(*
	FIFO queue that owns every FB_LogRecord pointer it contains. push drops the
	oldest owned records when the bound is reached. The bound is maxCount, but
	never more than TcOtlp_GVL.MAX_LOOP_COUNT: a maxCount of zero, or one above
	that limit, is held to MAX_LOOP_COUNT so that free always reaches the end.
	pop transfers ownership back to the caller. transferTo moves allocated
	nodes between queue owners without copying records.
*)
FUNCTION_BLOCK FB_LogRecordQueue
VAR
	_head: POINTER TO ST_LinkedListNode;
	_tail: POINTER TO ST_LinkedListNode;
	_cursor: POINTER TO ST_LinkedListNode;
END_VAR
VAR_OUTPUT
	count: UDINT;
	maxCount: UDINT;
	droppedCount: UDINT;
END_VAR

(* The enforced bound: maxCount, held to MAX_LOOP_COUNT when it is zero or larger. *)
METHOD _capacity : UDINT
IF THIS^.maxCount = 0 OR THIS^.maxCount > TcOtlp_GVL.MAX_LOOP_COUNT THEN
	_capacity := TcOtlp_GVL.MAX_LOOP_COUNT;
ELSE
	_capacity := THIS^.maxCount;
END_IF
END_METHOD

METHOD FB_Exit : BOOL
VAR_INPUT
	bInCopyCode: BOOL;
END_VAR
IF NOT bInCopyCode THEN
	THIS^.free();
END_IF
END_METHOD

METHOD FB_Init : BOOL
VAR_INPUT
	bInitRetains: BOOL;
	bInCopyCode: BOOL;
	maxCount: UDINT := 0;
END_VAR
THIS^.maxCount := maxCount;
END_METHOD

(*
	Releases every owned record. push holds count to MAX_LOOP_COUNT, so the loop
	always reaches the end. If it ever stops early, the unreleased nodes stay in
	the queue and free returns FALSE, so a later call can finish the job.
*)
METHOD free : BOOL
VAR
	_idx: UDINT;
	_node: POINTER TO ST_LinkedListNode;
	_record: POINTER TO FB_LogRecord;
END_VAR
FOR _idx := 0 TO TcOtlp_GVL.MAX_LOOP_COUNT DO
	IF THIS^._head = 0 THEN
		EXIT;
	END_IF

	_node := THIS^._head;
	THIS^._head := _node^.nxt;
	IF _node^.val <> 0 THEN
		_record := _node^.val;
		_node^.val := 0;
		_record^.delete(pSelf:=_record);
	END_IF
	__DELETE(_node);
	IF THIS^.count > 0 THEN
		THIS^.count := THIS^.count - 1;
	END_IF
END_FOR

THIS^._cursor := THIS^._head;
IF THIS^._head = 0 THEN
	THIS^._tail := 0;
	THIS^.count := 0;
END_IF
free := THIS^._head = 0;
END_METHOD

METHOD next : POINTER TO FB_LogRecord
next := 0;

IF THIS^._cursor <> 0 THEN
	next := THIS^._cursor^.val;
	THIS^._cursor := THIS^._cursor^.nxt;
END_IF
END_METHOD

METHOD pop : BOOL
VAR_IN_OUT
	pValue: POINTER TO FB_LogRecord;
END_VAR
VAR_OUTPUT
	failureReason: E_LogRecordQueueFailureReason;
END_VAR
VAR
	_node: POINTER TO ST_LinkedListNode;
END_VAR
pop := FALSE;
failureReason := E_LogRecordQueueFailureReason.NA;

IF pValue <> 0 THEN
	failureReason := E_LogRecordQueueFailureReason.DESTINATION_ALREADY_ASSIGNED;
	RETURN;
END_IF
IF THIS^._head = 0 THEN
	failureReason := E_LogRecordQueueFailureReason.QUEUE_EMPTY;
	RETURN;
END_IF

_node := THIS^._head;
THIS^._head := _node^.nxt;
IF THIS^._cursor = _node THEN
	THIS^._cursor := THIS^._head;
END_IF
IF THIS^._head = 0 THEN
	THIS^._tail := 0;
END_IF

pValue := _node^.val;
_node^.val := 0;
_node^.nxt := 0;
__DELETE(_node);
_node := 0;
THIS^.count := THIS^.count - 1;
pop := failureReason = E_LogRecordQueueFailureReason.NA;
END_METHOD

METHOD push : BOOL
VAR_IN_OUT
	pValue: POINTER TO FB_LogRecord;
END_VAR
VAR_OUTPUT
	failureReason: E_LogRecordQueueFailureReason;
END_VAR
VAR
	_node: POINTER TO ST_LinkedListNode;
	_droppedRecord: POINTER TO FB_LogRecord;
	_popFailureReason: E_LogRecordQueueFailureReason;
	_idx: UDINT;
	_bound: UDINT;
END_VAR
push := FALSE;
failureReason := E_LogRecordQueueFailureReason.NA;

IF pValue = 0 THEN
	failureReason := E_LogRecordQueueFailureReason.RECORD_POINTER_NULL;
	RETURN;
END_IF

// Allocate before evicting so an allocation failure leaves the queue unchanged.
_node := __NEW(ST_LinkedListNode);
IF _node = 0 THEN
	failureReason := E_LogRecordQueueFailureReason.MEMORY_ALLOCATION_FAILURE;
	RETURN;
END_IF

// maxCount is writable, so also restore the bound after a runtime reduction.
_bound := THIS^._capacity();
FOR _idx := 0 TO TcOtlp_GVL.MAX_LOOP_COUNT DO
	IF THIS^.count < _bound THEN
		EXIT;
	END_IF
	IF NOT THIS^.pop(pValue:=_droppedRecord, failureReason=>_popFailureReason) THEN
		__DELETE(_node);
		_node := 0;
		failureReason := _popFailureReason;
		RETURN;
	END_IF
	_droppedRecord^.delete(pSelf:=_droppedRecord);
	THIS^.droppedCount := THIS^.droppedCount + 1;
END_FOR
IF THIS^.count >= _bound THEN
	__DELETE(_node);
	_node := 0;
	failureReason := E_LogRecordQueueFailureReason.MAX_SIZE_ENFORCEMENT_FAILURE;
	RETURN;
END_IF

_node^.val := pValue;
_node^.nxt := 0;
IF THIS^._tail = 0 THEN
	THIS^._head := _node;
	THIS^._cursor := _node;
ELSE
	THIS^._tail^.nxt := _node;
END_IF
THIS^._tail := _node;
THIS^.count := THIS^.count + 1;
pValue := 0;
push := failureReason = E_LogRecordQueueFailureReason.NA;
END_METHOD

METHOD reset
THIS^._cursor := THIS^._head;
END_METHOD

(* Moves the head node to the tail without changing record ownership. *)
METHOD rotate : BOOL
VAR_OUTPUT
	failureReason: E_LogRecordQueueFailureReason;
END_VAR
VAR
	_node: POINTER TO ST_LinkedListNode;
END_VAR
rotate := FALSE;
failureReason := E_LogRecordQueueFailureReason.NA;

IF THIS^._head = 0 THEN
	failureReason := E_LogRecordQueueFailureReason.QUEUE_EMPTY;
	RETURN;
END_IF

IF THIS^._head <> THIS^._tail THEN
	_node := THIS^._head;
	THIS^._head := _node^.nxt;
	_node^.nxt := 0;
	THIS^._tail^.nxt := _node;
	THIS^._tail := _node;
END_IF

THIS^._cursor := THIS^._head;
rotate := failureReason = E_LogRecordQueueFailureReason.NA;
END_METHOD

(*
	Transfers the allocated nodes and owned records without copying them.
	The destination must be a different, empty queue. It receives up to count
	of the oldest records, also respecting the destination's bound.
*)
METHOD transferTo : BOOL
VAR_IN_OUT
	destination: FB_LogRecordQueue;
END_VAR
VAR_INPUT
	count: UDINT;
END_VAR
VAR_OUTPUT
	failureReason: E_LogRecordQueueFailureReason;
END_VAR
VAR
	_transferCount: UDINT;
	_idx: UDINT;
END_VAR
transferTo := FALSE;
failureReason := E_LogRecordQueueFailureReason.NA;

IF ADR(destination) = THIS THEN
	failureReason := E_LogRecordQueueFailureReason.SELF_TRANSFER_NOT_ALLOWED;
	RETURN;
END_IF
IF destination.count <> 0 OR_ELSE destination._head <> 0 OR_ELSE destination._tail <> 0 THEN
	failureReason := E_LogRecordQueueFailureReason.DESTINATION_NOT_EMPTY;
	RETURN;
END_IF

_transferCount := count;
IF _transferCount > THIS^.count THEN
	_transferCount := THIS^.count;
END_IF
IF _transferCount > destination._capacity() THEN
	_transferCount := destination._capacity();
END_IF
IF _transferCount = 0 THEN
	transferTo := failureReason = E_LogRecordQueueFailureReason.NA;
	RETURN;
END_IF

destination._head := THIS^._head;
destination._tail := destination._head;
FOR _idx := 1 TO _transferCount - 1 DO
	destination._tail := destination._tail^.nxt;
END_FOR

THIS^._head := destination._tail^.nxt;
destination._tail^.nxt := 0;
destination._cursor := destination._head;
destination.count := _transferCount;

THIS^.count := THIS^.count - _transferCount;
THIS^._cursor := THIS^._head;
IF THIS^._head = 0 THEN
	THIS^._tail := 0;
END_IF
transferTo := failureReason = E_LogRecordQueueFailureReason.NA;
END_METHOD

END_FUNCTION_BLOCK

(* stored: Version 1.1.0.1
   POU FB_LogRecordQueue: Id {9e1ecc03-058c-4b23-92d3-3bd422ae83cb}, SpecialFunc None
   Method _capacity: Id {29c1afd9-6ad2-4b61-af2f-13dab25e3140}
   Method FB_Exit: Id {6d9d65b6-2d68-47f0-b7cb-88e631d7acef}
   Method FB_Init: Id {c957bb4c-b6fd-49dc-a4b2-5cb85e435a28}
   Method free: Id {fbd1c94b-c09e-4d95-a598-0cd5bb8a61f6}
   Method next: Id {720ec83f-b785-4449-92d1-d6ec1cfa78ab}
   Method pop: Id {81f42449-d168-4086-9f3b-beae690752ef}
   Method push: Id {160c78e0-3b3f-49cd-8c42-eefe5336e9d8}
   Method reset: Id {8e5c6da1-a3e7-4711-8032-291e4a16dc6e}
   Method rotate: Id {38f6dc88-7df0-47e8-9ca7-d6d6b143b68e}
   Method transferTo: Id {e7eb4308-b34a-4dc8-852c-97a5624b88e2} *)
